Fanuc KAREL source: kb00050.KL

-- PROVISIONAL review KL for V940-1; original PC SHA256 a191d7731de3193f2545652319c9eb03574314a114e5bbb6fbed71638e2fda77
-- Incomplete behavior may be omitted. Consult companion uncertainty JSON. Do not deploy.
PROGRAM KB00050
%NOLOCKGROUP
BEGIN
  -- V9_ZERO_TABLE_METADATA_HINT layout=0002_ascii; no indexed target words; source/name/runtime held
  -- UNRESOLVED_PC offsets 5-14; opcodes 3F,75
  -- UNRESOLVED_PC offsets 19-28; opcodes 3F,75
  -- UNRESOLVED_PC offsets 33-42; opcodes 3F,75
  -- UNRESOLVED_PC offsets 47-56; opcodes 3F,75
  -- UNRESOLVED_PC offsets 61-68; opcodes 9D,23
  -- UNRESOLVED_PC offsets 73-80; opcodes 9D,23
  -- UNRESOLVED_PC offsets 85-92; opcodes 9D,23
  -- UNRESOLVED_PC offsets 97-104; opcodes 9D,23
  -- UNRESOLVED_PC offsets 109-116; opcodes 9D,23
  -- UNRESOLVED_PC offsets 121-189; opcodes 27,22,2A,22,2A,22,2A,22,2A,22,22,22,22,22,27,9D,31
  -- UNRESOLVED_PC offsets 194-198; opcodes 7F
END KB00050
